TYPE tea :
STRUCT

Name			: STRING;
Price			: REAL;
ingredients		: STRING;	


END_STRUCT
END_TYPE

(* stored: Version 1.1.0.1
   DUT tea: Id {3deb03eb-6095-44ca-85a3-1787ae1f3249} *)
